Fanuc KAREL source: ko00083.KL

-- PROVISIONAL review KL for V770-1; original PC SHA256 a9e9ca48a413476e1716234fbe2b61c5ed36ffd42eea2f7a4d6e965053d61482
-- Incomplete behavior may be omitted. Consult companion uncertainty JSON. Do not deploy.
PROGRAM KO00083
%NOLOCKGROUP
BEGIN
  -- UNRESOLVED_PC offsets 5-12; opcodes 9D,23
  -- UNRESOLVED_PC offsets 17-66; opcodes 27,27,49,7E,AD,22,1C,22,31,7E,4A
  -- UNRESOLVED_PC offsets 71-75; opcodes 7F
END KO00083
